// TIA Portal V20 export
// export: Created 2026-10-19T18:36:46.8242776Z, ExportSetting WithDefaults, DisplayName Totally Integrated Automation Portal, DisplayVersion V20 Update 6, DisplayName TIA Portal Openness, DisplayVersion V20 Update 6, DisplayName TIA Portal Version Control Interface, DisplayVersion V20 Update 6, DisplayName SINAMICS Startdrive Advanced, DisplayVersion V20 SP1, DisplayName SINAMICS Startdrive G130, G150, S120, S150, SINAMICS MV, G220, S200, S210, DisplayVersion V20 SP1, DisplayName SINAMICS Startdrive G110M, G120, G120C, G120D, G120P, G115D, DisplayVersion V20 SP1, DisplayName STEP 7 Professional, DisplayVersion V20 Update 6, DisplayName STEP 7 Safety, DisplayVersion V20 Update 2, DisplayName WinCC Basic/Comfort/Advanced, DisplayVersion V20 Update 6, DisplayName WinCC Unified, DisplayVersion V20 Update 6
FUNCTION "OT_Charge_Commands" : Void   // FC52, SCL
{ S7_Optimized_Access := 'TRUE' }
VERSION : 0.1
// stored: AutoNumber true, IsIECCheckEnabled false, SetENOAutomatically false, UDAEnableTagReadback false
   VAR_IN_OUT
      Auto_Test : "Auto_Test";
   END_VAR
BEGIN
   "OrderTable_HMI"."Manual order" := #Auto_Test.Manual;
   "OrderTable_HMI"."From level" := #Auto_Test."From level";
   "OrderTable_HMI"."To level" := #Auto_Test."To level";
   "OrderTable_HMI"."Testing Time" := #Auto_Test."Testing Time";
   "OrderTable_HMI"."Numer of cycles" := #Auto_Test."Numer of cycles";
   "OrderTable_HMI".Level := UINT_TO_BYTE(#Auto_Test.Level);
END_FUNCTION
